// TIA Portal V20 export
// export: Created 2026-10-12T15:46:51.3857994Z, ExportSetting WithDefaults, DisplayName Totally Integrated Automation Portal, DisplayVersion V20, DisplayName TIA Portal Openness, DisplayVersion V20, DisplayName TIA Portal Teamcenter Gateway, DisplayVersion V20, DisplayName TIA Portal Version Control Interface, DisplayVersion V20, DisplayName SINAMICS Startdrive Advanced, DisplayVersion V20 SP1 Update 2, DisplayName SINAMICS Startdrive G110M, G120, G120C, G120D, G120P, G115D, DisplayVersion V20 SP1 Update 2, DisplayName SINAMICS Startdrive G130, G150, S120, S150, SINAMICS MV, G220, S200, S210, DisplayVersion V20 SP1 Update 2, DisplayName STEP 7 Professional, DisplayVersion V20, DisplayName STEP 7 Safety, DisplayVersion V20, DisplayName WinCC Basic/Comfort/Advanced, DisplayVersion V20, DisplayName WinCC Professional, DisplayVersion V20, DisplayName WinCC Unified, DisplayVersion V20
FUNCTION "FRK_JsonPut" : Bool   // FC116, SCL
{ S7_Optimized_Access := 'TRUE' }
VERSION : 0.1
// Append complete text or refuse. Explicit destination width and length check
//  protect long WSTRING lines against truncation in the Siemens string runtime.
// stored: AutoNumber true, IsIECCheckEnabled false, SetENOAutomatically false, UDAEnableTagReadback false
   VAR_INPUT
      Text : WString;
   END_VAR
   VAR_IN_OUT
      Line : WString;
   END_VAR
   VAR_TEMP
      Expected : Int;
   END_VAR
BEGIN

   #FRK_JsonPut := FALSE;
   #Expected := LEN(#Line) + LEN(#Text);
   IF #Expected > 480 THEN
       RETURN;
   END_IF;
   #Line := CONCAT(IN1 := #Line, IN2 := #Text);
   #FRK_JsonPut := LEN(#Line) = #Expected;
END_FUNCTION
